PROGRAM Axis_test
VAR
    // Online commands: bMoveAbsolute and bStop are rising-edge commands.
    bPower : BOOL := FALSE;
    bMoveAbsolute : BOOL := FALSE;
    bStop : BOOL := FALSE;
	bReset : BOOL := FALSE;

    // Values use the engineering unit configured for the selected NC axis.
    lrTargetPosition : LREAL := 0.0;
    lrVelocity : LREAL := 5.0;
    lrAcceleration : LREAL := 20.0;
    lrDeceleration : LREAL := 20.0;
    lrJerk : LREAL := 100.0;

    // Online diagnostics.
    bPowerStatus : BOOL;
    bMoveBusy : BOOL;
    bMoveDone : BOOL;
    bStopDone : BOOL;
    bError : BOOL;
    udiErrorID : UDINT;
    lrActualPosition : LREAL;

    fbAxisTest : FB_AxisPositionTest;
END_VAR

fbAxisTest(
    bPower := bPower,
    bMoveAbsolute := bMoveAbsolute,
	bReset := bReset,
    bStop := bStop,
    lrTargetPosition := lrTargetPosition,
    lrVelocity := lrVelocity,
    lrAcceleration := lrAcceleration,
    lrDeceleration := lrDeceleration,
    lrJerk := lrJerk,
    // Change only this line to select another test axis.
    Axis := GVL_Motion.gAxisConveyor,
    bPowerStatus => bPowerStatus,
    bMoveBusy => bMoveBusy,
    bMoveDone => bMoveDone,
    bStopDone => bStopDone,
    bError => bError,
    udiErrorID => udiErrorID,
    lrActualPosition => lrActualPosition);

END_PROGRAM

(* stored: Version 1.1.0.1, ProductVersion 3.1.4024.16
   POU Axis_test: Id {f0a9d9de-a053-4cc5-a6aa-b4563593a597}, SpecialFunc None *)
